Fanuc KAREL source: kt00407.KL

-- PROVISIONAL review KL for V1013-1; original PC SHA256 e7a953310ebb1cdf29ef30bb052f43ee57bacd86672f7b1e6a84db5fc9111900
-- Incomplete behavior may be omitted. Consult companion uncertainty JSON. Do not deploy.
PROGRAM KT00407
%NOLOCKGROUP
VAR
  R1 : REAL
  OUT : BOOLEAN
-- UNRESOLVED_DECL Y2 type=002018
BEGIN
  -- UNRESOLVED_PC offsets 5-16; opcodes 2E,23
  -- UNRESOLVED_PC offsets 21-35; opcodes 2E,22,9D,33,B2
  -- UNRESOLVED_PC offsets 40-63; opcodes 21,22,9D,33,B1,64,71,23
  -- UNRESOLVED_PC offsets 68-72; opcodes 7F
END KT00407
